(* IEC 61131-3 sources: nautilus/examples/lift-station, 3 files *)

(* ---- field_map.st ---- *)
PROGRAM FieldMap
(* Field-only tag glue — the one place this project departs from "the same
   program files run on the bench and in the field." `naut modbus import`
   names every tag `<instance-id>_<register-tag>` unconditionally (see
   modbus/codegen/devicemap.go); there is no way to suppress the prefix,
   so a bare name like `LSHH101` cannot come out of ANY instance id, and
   `P101`/`P102` are already spoken for by the VFD instances, so the RIO's
   seal-fail/over-temp points can't reuse them either. The RIO instance
   (devices.yaml, id RIO) therefore imports as RIO_Level, RIO_Flow,
   RIO_LSHH101, RIO_LSLL101, RIO_P101_SealFail, RIO_P101_OverTemp,
   RIO_P102_SealFail, RIO_P102_OverTemp — and this task, which only exists
   in field.yaml, renames them onto the canonical tags every other program
   (sequence.sfc, level.fbd, permissives.ld, stats.st) actually reads: the
   same names the bench manifest's sim task writes directly. Logged in
   docs/design/examples-dogfood.md. *)
VAR_EXTERNAL
    RIO_Level         : REAL;
    RIO_Flow          : REAL;
    RIO_LSHH101       : BOOL;
    RIO_LSLL101       : BOOL;
    RIO_P101_SealFail : BOOL;
    RIO_P101_OverTemp : BOOL;
    RIO_P102_SealFail : BOOL;
    RIO_P102_OverTemp : BOOL;

    LIT101_Level  : REAL;
    FIT101_Flow   : REAL;
    LSHH101       : BOOL;
    LSLL101       : BOOL;
    P101_SealFail : BOOL;
    P101_OverTemp : BOOL;
    P102_SealFail : BOOL;
    P102_OverTemp : BOOL;
END_VAR
LIT101_Level  := RIO_Level;
FIT101_Flow   := RIO_Flow;
LSHH101       := RIO_LSHH101;
LSLL101       := RIO_LSLL101;
P101_SealFail := RIO_P101_SealFail;
P101_OverTemp := RIO_P101_OverTemp;
P102_SealFail := RIO_P102_SealFail;
P102_OverTemp := RIO_P102_OverTemp;
END_PROGRAM

(* ---- sim.st ---- *)
PROGRAM WetWell
(* Bench-only plant: WW-101 (level from an inflow/outflow balance, via
   lib/physics.st's WetWellModel) and two submersible-pump/VFD models
   (VfdModel). Inflow is InflowGpm plus a slow sinusoid (+-20 %) so the
   level never sits dead flat; InflowGpm set to 950 is the "storm" the
   design calls out. A real deployment deletes this task entirely —
   field.yaml has no sim task and points the same control programs at
   the real devices instead (see docs/design/examples-dogfood.md for the
   one place the field tag names needed a small glue program). *)
VAR_EXTERNAL
    LIT101_Level : REAL;
    LSHH101      : BOOL;
    LSLL101      : BOOL;
    FIT101_Flow  : REAL;
    SimDtS       : REAL;
    InflowGpm    : REAL;
    ForceLSHH    : BOOL;

    P101_RunCmd      : BOOL;
    P101_SpeedCmd    : REAL;
    P101_Running     : BOOL;
    P101_SpeedHz     : REAL;
    P101_Amps        : REAL;
    P101_VfdFault    : BOOL;
    P101_InjectFault : BOOL;
    P101_SealFail        : BOOL;
    P101_InjectSealFail  : BOOL;
    P101_OverTemp        : BOOL;
    P101_InjectOverTemp  : BOOL;
    P101_FlapOverTemp    : BOOL;

    P102_RunCmd      : BOOL;
    P102_SpeedCmd    : REAL;
    P102_Running     : BOOL;
    P102_SpeedHz     : REAL;
    P102_Amps        : REAL;
    P102_VfdFault    : BOOL;
    P102_InjectFault : BOOL;
    P102_SealFail        : BOOL;
    P102_InjectSealFail  : BOOL;
    P102_OverTemp        : BOOL;
    P102_InjectOverTemp  : BOOL;
END_VAR
VAR
    well   : WetWellModel;
    vfd101 : VfdModel;
    vfd102 : VfdModel;
    tSec   : REAL;
    flapS  : REAL;
END_VAR
VAR CONSTANT
    InflowVaryFrac : REAL := 0.20;
    InflowPeriodS  : REAL := 240.0;
    TwoPi          : REAL := 6.2831853;
END_VAR

tSec := tSec + SimDtS;

vfd101(RunCmd := P101_RunCmd, SpeedCmd := P101_SpeedCmd, Dt := SimDtS, InjectFault := P101_InjectFault,
       Running => P101_Running, SpeedHz => P101_SpeedHz, Amps => P101_Amps, Fault => P101_VfdFault);
vfd102(RunCmd := P102_RunCmd, SpeedCmd := P102_SpeedCmd, Dt := SimDtS, InjectFault := P102_InjectFault,
       Running => P102_Running, SpeedHz => P102_SpeedHz, Amps => P102_Amps, Fault => P102_VfdFault);

(* Seal-leak and over-temp probes have no physics to speak of: pass the
   bench inject tags straight through, exactly like a wire from a switch. *)
P101_SealFail := P101_InjectSealFail;
(* A contact that chatters: with the flap tag set, P-101's over-temp probe is
   made for 3 s and broken for 2 s, over and over, the way a marginal
   contact or a hunting thermostat does. The alarm's 2 s on-delay lets
   each 3 s make through, so it activates every 5 s: chatter within a
   minute. Bench only. *)
flapS := flapS + SimDtS;
IF flapS >= 5.0 THEN
    flapS := 0.0;
END_IF;
P101_OverTemp := P101_InjectOverTemp OR (P101_FlapOverTemp AND flapS < 3.0);
P102_SealFail := P102_InjectSealFail;
P102_OverTemp := P102_InjectOverTemp;

FIT101_Flow := PumpFlowGpm(P101_SpeedHz) + PumpFlowGpm(P102_SpeedHz);

well(InflowGpm := InflowGpm * (1.0 + InflowVaryFrac * SIN(tSec / InflowPeriodS * TwoPi)),
     OutflowGpm := FIT101_Flow, Dt := SimDtS, Level := LIT101_Level);

(* The floats switch with a differential, as a real tilt float does: it
   trips at one level and resets a few inches past it, so a level sitting
   on the mark doesn't make it chatter. *)
IF ForceLSHH THEN
    LSHH101 := TRUE;
ELSIF LIT101_Level >= 95.0 THEN
    LSHH101 := TRUE;
ELSIF LIT101_Level <= 91.0 THEN
    LSHH101 := FALSE;
END_IF;
IF LIT101_Level <= 8.0 THEN
    LSLL101 := TRUE;
ELSIF LIT101_Level >= 12.0 THEN
    LSLL101 := FALSE;
END_IF;
END_PROGRAM

(* ---- stats.st ---- *)
PROGRAM Stats
(* Runtime hours/starts for each pump (RuntimeMeter, lib/pump.st) and the
   station flow totalizer. Shared, unchanged, between the bench and field
   manifests — it only reads process values and writes rollups, never a
   role that differs between them. *)
VAR_EXTERNAL
    P101_Running : BOOL;
    P102_Running : BOOL;
    P101_Stats   : PumpStats;
    P102_Stats   : PumpStats;
    FIT101_Flow  : REAL;
    StationFlowGal: REAL;
    StatsDtS     : REAL;
END_VAR
VAR
    meter101 : RuntimeMeter;
    meter102 : RuntimeMeter;
END_VAR
meter101(Running := P101_Running, Dt := StatsDtS, Stats := P101_Stats);
meter102(Running := P102_Running, Dt := StatsDtS, Stats := P102_Stats);

(* Totalized discharge volume, gal: gal/min * s / 60. *)
StationFlowGal := StationFlowGal + FIT101_Flow * StatsDtS / 60.0;
END_PROGRAM
